Staubli VAL3: insertCirclePoint.pgx

public program insertCirclePoint(string x_sKey, num x_nIndex, bool& x_bToSave)
  local num l_j
  local frame l_fFrame
  local tool l_tTool
  local num l_i
  local num l_nFrameIndex
  local num l_nToolIndex
  local pointRx l_pPoint
begin
  //  link(l_fFrame,world)
  //  link(l_tTool,flange)
  //  call savedata:getFrame(trajTemp:tTrajItem[x_sKey].nFrameIndex,l_fFrame)
  //  call savedata:getTool(trajTemp:tTrajItem[x_sKey].nToolIndex,l_tTool)
  //insert(trajTemp:tTrajItem[x_sKey].pPointItem[x_nIndex+1])
  append(trajTemp:tTrajItem[x_sKey].pPointItem)

  for l_i = (size(trajTemp:tTrajItem[x_sKey].pPointItem)-1) to(x_nIndex+1) step -1
    //logMsg(toString("",l_i))
    call copyPoint3(x_sKey,l_i,l_i-1)
  endFor
  //2024.12.06 当前位置作为插入点坐标
  l_nFrameIndex=trajTemp:tTrajItem[x_sKey].nFrameIndex
  l_nToolIndex=trajTemp:tTrajItem[x_sKey].nToolIndex
  call savedata:getFrame(l_nFrameIndex,l_fFrame)
  call savedata:getTool(l_nToolIndex,l_tTool)
  trajTemp:tTrajItem[x_sKey].pPointItem[x_nIndex+1].jJointRx=herej()
  l_pPoint=jointToPoint(l_tTool,l_fFrame,herej())
  trajTemp:tTrajItem[x_sKey].pPointItem[x_nIndex+1].pPointRx.trsf=l_pPoint.trsf
  trajTemp:tTrajItem[x_sKey].pPointItem[x_nIndex+1].pPointRx.config=l_pPoint.config
  trajTemp:tTrajItem[x_sKey].pPointItem[x_nIndex+1].pInter.trsf=l_pPoint.trsf
  trajTemp:tTrajItem[x_sKey].pPointItem[x_nIndex+1].pInter.config=l_pPoint.config
  //

  //trajTemp:tTrajItem[x_sKey].pPointItem[x_nIndex+1].pPointRx=trajTemp:tTrajItem[x_sKey].pPointItem[x_nIndex].pPointRx
  //trajTemp:tTrajItem[x_sKey].pPointItem[x_nIndex+1].jJointRx=trajTemp:tTrajItem[x_sKey].pPointItem[x_nIndex].jJointRx
  trajTemp:tTrajItem[x_sKey].pPointItem[x_nIndex+1].pParaItem.mMdesc=trajTemp:tTrajItem[x_sKey].pPointItem[x_nIndex].pParaItem.mMdesc
  trajTemp:tTrajItem[x_sKey].pPointItem[x_nIndex+1].pParaItem.nMoveType=2
  trajTemp:tTrajItem[x_sKey].pPointItem[x_nIndex+1].pParaItem.nDelay=trajTemp:tTrajItem[x_sKey].pPointItem[x_nIndex].pParaItem.nDelay
  trajTemp:tTrajItem[x_sKey].pPointItem[x_nIndex+1].pParaItem.nSigValue=trajTemp:tTrajItem[x_sKey].pPointItem[x_nIndex].pParaItem.nSigValue
  trajTemp:tTrajItem[x_sKey].pPointItem[x_nIndex+1].pParaItem.nActionIndex=trajTemp:tTrajItem[x_sKey].pPointItem[x_nIndex].pParaItem.nActionIndex
  trajTemp:tTrajItem[x_sKey].pPointItem[x_nIndex+1].pParaItem.nPercentage=trajTemp:tTrajItem[x_sKey].pPointItem[x_nIndex].pParaItem.nPercentage
  for l_j = 0 to 2
    trajTemp:tTrajItem[x_sKey].pPointItem[x_nIndex+1].pParaItem.iIfItem.nSigType[l_j]=trajTemp:tTrajItem[x_sKey].pPointItem[x_nIndex].pParaItem.iIfItem.nSigType[l_j]
    trajTemp:tTrajItem[x_sKey].pPointItem[x_nIndex+1].pParaItem.iIfItem.nSigIndex[l_j]=trajTemp:tTrajItem[x_sKey].pPointItem[x_nIndex].pParaItem.iIfItem.nSigIndex[l_j]
    trajTemp:tTrajItem[x_sKey].pPointItem[x_nIndex+1].pParaItem.iIfItem.nValue[l_j]=trajTemp:tTrajItem[x_sKey].pPointItem[x_nIndex].pParaItem.iIfItem.nValue[l_j]
  endFor
  //trajTemp:libSave()
  x_bToSave=true
end
